FUNCTION_BLOCK "TiaMcpLibraryGate"
{ S7_Optimized_Access := 'TRUE' }
VERSION : 0.1
VAR_INPUT
    Enable : Bool;
END_VAR
VAR_OUTPUT
    Ready : Bool;
END_VAR
BEGIN
    #Ready := NOT #Enable;
END_FUNCTION_BLOCK
